SUBAPPLICATION AULI_GT_0 (* Prüft ob ULINT-Adapter Wert > 0 ist (AX-Adapter Ausgang) *)
  (* Standard: 61499-2 *)
  (* Version 1.0, 2026-10-15, franz, Meisterschulen am Ostbahnhof *)
  PACKAGE MyLib::sys;
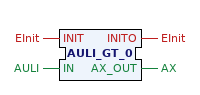
  EVENT_INPUT
    INIT : EInit; (* Initialization Request *)
  END_EVENT
  EVENT_OUTPUT
    INITO : EInit; (* Initialization Confirm *)
  END_EVENT
  SOCKETS
    IN : adapter::types::unidirectional::AULI;
  END_SOCKETS
  PLUGS
    AX_OUT : adapter::types::unidirectional::AX;
  END_PLUGS
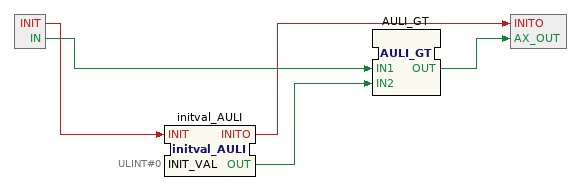
  FBS
    AULI_GT : adapter::iec61131::comparison::AULI_GT;
    initval_AULI : adapter::types::unidirectional::AULI::initval::initval_AULI(INIT_VAL := ULINT#0);
  END_FBS
  EVENT_CONNECTIONS
    INIT TO initval_AULI.INIT;
    initval_AULI.INITO TO INITO;
  END_CONNECTIONS
  ADAPTER_CONNECTIONS
    IN TO AULI_GT.IN1;
    AULI_GT.OUT TO AX_OUT;
    initval_AULI.OUT TO AULI_GT.IN2;
  END_CONNECTIONS
END_SUBAPPLICATION
